FUNCTION_BLOCK Panel_button_cotrol (* Basic Function Block Type *)
  (* Standard: 61499-2 *)
  (* Version 0.0, 10/19/2026, lizar, Schneider Electric, Template *)
  PACKAGE Main;
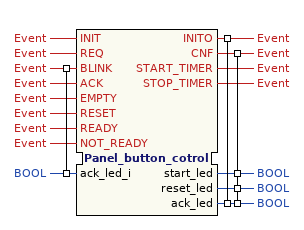
  EVENT_INPUT
    INIT; (* Initialization Request *)
    REQ; (* Normal Execution Request *)
    BLINK WITH ack_led_i;
    ACK;
    EMPTY;
    RESET;
    READY;
    NOT_READY;
  END_EVENT
  EVENT_OUTPUT
    INITO WITH ack_led; (* Initialization Confirm *)
    CNF WITH ack_led, start_led, reset_led; (* Execution Confirmation *)
    START_TIMER;
    STOP_TIMER;
  END_EVENT
  VAR_INPUT
    ack_led_i : BOOL;
  END_VAR
  VAR_OUTPUT
    start_led : BOOL;
    reset_led : BOOL;
    ack_led : BOOL; (* Output event qualifier *)
  END_VAR
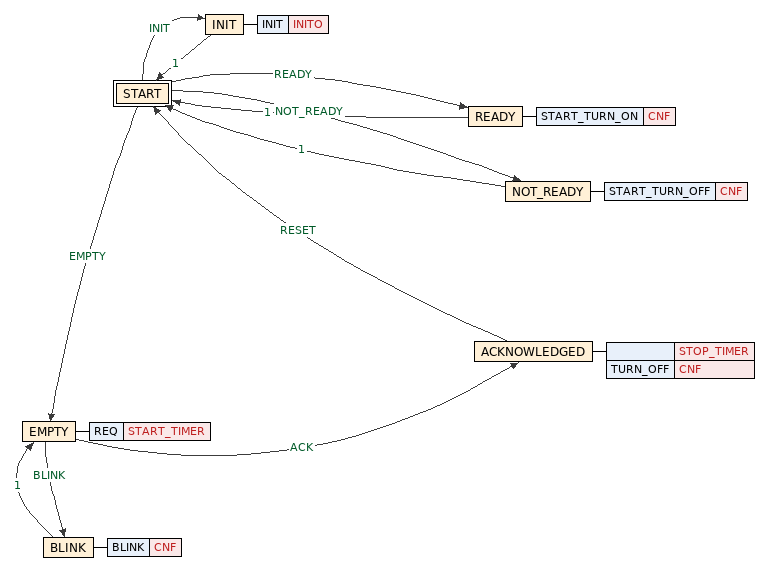
  EC_STATES
    START; (* Initial State *)
    INIT : INIT -> INITO; (* Initialization *)
    EMPTY : REQ -> START_TIMER; (* Normal execution *)
    BLINK : BLINK -> CNF;
    ACKNOWLEDGED : -> STOP_TIMER, TURN_OFF -> CNF;
    READY : START_TURN_ON -> CNF;
    NOT_READY : START_TURN_OFF -> CNF;
  END_STATES
  EC_TRANSITIONS
    START TO INIT := INIT;
    INIT TO START := 1;
    EMPTY TO BLINK := BLINK;
    BLINK TO EMPTY := 1;
    EMPTY TO ACKNOWLEDGED := ACK;
    ACKNOWLEDGED TO START := RESET;
    START TO READY := READY;
    READY TO START := 1;
    START TO EMPTY := EMPTY;
    START TO NOT_READY := NOT_READY;
    NOT_READY TO START := 1;
  END_TRANSITIONS
  ALGORITHM INIT IN ST: (* Initialization algorithm *)
;
ack_led:=TRUE;
  END_ALGORITHM
  ALGORITHM REQ IN ST: (* Normally executed algorithm *)
;
  END_ALGORITHM
  ALGORITHM BLINK IN ST:
;
ack_led := NOT(ack_led_i);
  END_ALGORITHM
  ALGORITHM TURN_OFF IN ST:
;
ack_led:=FALSE;
  END_ALGORITHM
  ALGORITHM START_TURN_ON IN ST:
;
start_led:=TRUE;
  END_ALGORITHM
  ALGORITHM START_TURN_OFF IN ST:
;

start_led:=FALSE;
  END_ALGORITHM
END_FUNCTION_BLOCK
